(* Logix 5000 project; controller AOI_Working vendor 1 type 14 code 166 rev 35.11; software revision 35.04 *)

TASK MainTask (continuous, watchdog 500 ms) : MainProgram
TASK Normal_500ms (periodic, rate 500 ms, priority 10, watchdog 500 ms) : Main

MODULES
   Local : vendor 1 type 14 code 166 (ICP 0, rev 35.11)
END_MODULES

ADD_ON_INSTRUCTION AnalogInput   (* revision 1.1, vendor NixSoftware *)
// Simple scaling routine for analog inputs.
// Converts between raw units to EU
VAR_INPUT
   Inp_PVRaw : REAL; {required}   // Raw Input from I/O Point
   Cfg_InpRawMax : REAL := 100.0; {visible}   // Raw Value - Maximum Reading (Used for Scaling)
   Cfg_InpRawMin : REAL; {visible}   // Raw Value - Minimum Reading (Used for Scaling)
   Cfg_PVEUMax : REAL := 100.0; {visible}   // PV Maximum Value (In Engineering Units)
   Cfg_PVEUMin : REAL; {visible}   // PV Minimum Value (In Engineering Units)
END_VAR
VAR_OUTPUT
   Val_PV : REAL; {visible}   // Scaled PV (EU)
END_VAR
VAR_INPUT
   Sts_RangeError : BOOL;   // 1 = Range Invalid, Check Max/Mins
   Sts_CfgError : BOOL;   // 1 = Check Range, Protects against dividing by 0
END_VAR
VAR
   HMI_IOAssignment : STRING; {access None}
   HMI_Description : STRING; {access None}
   HMI_DisplayTag : STRING; {access None}
   _EUSpan : REAL; {access None}
   _RawSpan : REAL; {access None}
END_VAR

ROUTINE Logic   (* structured text *)
// Simple scaling routine for analog inputs.
// Converts between raw units to EU
   (* ============================================================
      Analog Input Scaling - Engineering Units Conversion
      Project  : Inavant Custom AOI Library
      AOI Name : AnalogInput
      ============================================================ *)
   
   (* --- Parameters / Tags (map to AOI InOut or UDT members) ---
      Inp_PVRaw       : REAL  - Raw analog input value (e.g. 0.0–32767.0 or 4.0–20.0 mA)
      Cfg_InpRawMin   : REAL  - Raw value corresponding to engineering minimum (e.g. 0.0 or 4.0)
      Cfg_InpRawMax   : REAL  - Raw value corresponding to engineering maximum (e.g. 32767.0 or 20.0)
      Cfg_EUMin       : REAL  - Engineering unit minimum (e.g. 0.0 PSI)
      Cfg_EUMax       : REAL  - Engineering unit maximum (e.g. 100.0 PSI)
      Val_PV         : REAL   - Scaled output in engineering units
      Sts_RangeErr    : BOOL  - Fault bit: TRUE if raw input is out of configured range
      Sts_DivZeroFlt  : BOOL  - Fault bit: TRUE if raw span is zero (invalid config)
   *)
   (* --- Clear faults from previous scan --- *)
   Sts_CfgError 		:= 0;
   Sts_RangeError   	:= 0;
   
   (* --- Guard: detect zero-span configuration --- *)
   _RawSpan := Cfg_InpRawMax - Cfg_InpRawMin;
   
   IF _RawSpan = 0.0 THEN
       (* Invalid config — cannot divide by zero; hold last good output *)
       Sts_CfgError := 1;
   
   ELSE
       (* --- Range check (informational, does NOT clamp output) --- *)
       IF (Inp_PVRaw < Cfg_InpRawMin) OR (Inp_PVRaw > Cfg_InpRawMax) THEN
           Sts_RangeError := 1;
       END_IF;
       (* --- Scaling equation --- *)
       Val_PV  := (Inp_PVRaw - Cfg_InpRawMin) * ((Cfg_PVEUMax - Cfg_PVEUMin) / (Cfg_InpRawMax - Cfg_InpRawMin)) + Cfg_PVEUMin;
   END_IF;
END_ROUTINE
END_ADD_ON_INSTRUCTION

ADD_ON_INSTRUCTION Inv_AI   (* revision 1.1, vendor NixSoftware *)
// Used for scaling a raw analog value to engineering units, includes alarm statuses and debounces.
VAR_INPUT
   Inp_PV : REAL; {visible}
   Inp_IOStatus : BOOL := 1; {visible}   // 1 = I/O Status is Good 0 = Alarm, generates Sts_Fail
   Inp_LoLoGate : BOOL := 1; {visible}   // 1 = Low-Low Sts Enabled
   Inp_LoGate : BOOL := 1; {visible}   // 1 = Low Sts Enabled
   Inp_HiGate : BOOL := 1; {visible}   // 1 = High Sts Enabled
   Inp_HiHiGate : BOOL := 1; {visible}   // 1 = High-High Sts Enabled
   Inp_FailGate : BOOL := 1; {visible}   // 1 = Fail Sts Enabled
   Cfg_InpRawMin : REAL; {visible}
   Cfg_InpRawMax : REAL := 100.0; {visible}
   Cfg_PVEUMin : REAL; {visible}
   Cfg_PVEUMax : REAL := 100.0; {visible}
   Cfg_HiHiLim : REAL := 1.5e+20;
   Cfg_HiHiDB : REAL := 1.0;
   Cfg_HiLim : REAL := 1.5e+20;
   Cfg_HiDB : REAL := 1.0;
   Cfg_LoLim : REAL := -1.5e+20;
   Cfg_LoDB : REAL := 1.0;
   Cfg_LoLoLim : REAL := -1.5e+20;
   Cfg_LoLoDB : REAL := 1.0;
   Cfg_FailHiLim : REAL := 104.0;   // PV (EU) High Fail Limit
   Cfg_FailLoLim : REAL := -3.0;   // PV (EU) Low Fail Limit
   Cfg_FailDB : REAL := 0.5;   // Failed PV DB
   Cfg_HiHiDlyOn : ALIAS FOR HiHi_Debounce.Cfg_DebounceON; {access None}
   Cfg_HiHiDlyOff : ALIAS FOR HiHi_Debounce.Cfg_DebounceOFF; {access None}
   Cfg_HiDlyOn : ALIAS FOR Hi_Debounce.Cfg_DebounceON; {access None}
   Cfg_HiDlyOff : ALIAS FOR Hi_Debounce.Cfg_DebounceOFF; {access None}
   Cfg_LoDlyOn : ALIAS FOR Lo_Debounce.Cfg_DebounceON; {access None}
   Cfg_LoDlyOff : ALIAS FOR Lo_Debounce.Cfg_DebounceOFF; {access None}
   Cfg_LoLoDlyOn : ALIAS FOR LoLo_Debounce.Cfg_DebounceON; {access None}
   Cfg_LoLoDlyOff : ALIAS FOR LoLo_Debounce.Cfg_DebounceOFF; {access None}
   Cfg_FailDlyOn : ALIAS FOR Fail_Debounce.Cfg_DebounceON; {access None}
   Cfg_FailDlyOff : ALIAS FOR Fail_Debounce.Cfg_DebounceOFF; {access None}
   Cfg_PVDecPlcs : INT := 2;
   Cfg_FiltTC : REAL;
END_VAR
VAR_OUTPUT
   Val : REAL; {access Read Only, visible}   // PV (EU)
   Sts_HiHi : BOOL; {visible}   // 1 = High-High Alarm Active
   Sts_Hi : BOOL; {visible}   // 1 = High Alarm Active
   Sts_Lo : BOOL; {visible}   // 1 = Low Alarm Active
   Sts_LoLo : BOOL; {visible}   // 1 = Low-Low Alarm Active
   Sts_Err : BOOL; {access Read Only, visible}   // 1 = Error in Configuration
   Sts_Fail : BOOL; {access Read Only, visible}   // 1 = Failed PV (Out of Range)
   Sts_FaultPresent : BOOL; {access Read Only}
   Val_Fault : DINT; {access Read Only}   // 0 = None 1 = Low Alm 2 = Hi Alm 3 = LoLo Alm 4 = HiHi Alm 32 = Failed PV 34 = Config. Error
   Val_PVEUMax : REAL; {access None, visible}
   Val_PVEUMin : REAL; {access None, visible}
END_VAR
VAR
   HMI_EU : STRING; {access None}
   HMI_Description : STRING; {access None}
   HMI_DisplayTag : STRING; {access None}
   HMI_Rack : STRING := 'RXXX'; {access None}
   HMI_Slot : STRING := 'SXX'; {access None}
   HMI_Channel : STRING := 'Ch.XX'; {access None}
   Wrk_InpDINT : DINT; {access None}
   Wrk_InpInfNaN : BOOL; {access None}
   Wrk_CalcedPV : REAL; {access None}   // Scaled Value - Pre Filtering
   Wrk_ScanT : TIMER := (PRE := 2147483647); {access None}
   HiHi_Debounce : Inv_Debounce; {access None}   // HiHi Alarm Debounce
   Wrk_HiHi : BOOL; {access None}   // Internal flag: High-High Status
   Hi_Debounce : Inv_Debounce; {access None}   // High Alarm Debounce
   Wrk_Hi : BOOL; {access None}   // Internal flag: High Status
   Wrk_Lo : BOOL; {access None}   // Internal flag: Lo Status
   Lo_Debounce : Inv_Debounce; {access None}   // Low Alarm Debounce
   Wrk_LoLo : BOOL; {access None}   // Internal Flag: Low-Low Status
   LoLo_Debounce : Inv_Debounce; {access None}   // Low-Low Alarm Debounce
   Wrk_Fault : DINT; {access None}   // Internal Fault Monitoring Tag
   Wrk_Fail : BOOL; {access None}   // Internal Flag: Fail Status
   Fail_Debounce : Inv_Debounce; {access None}   // Fail Alarm Debounce
   Wrk_Alpha : REAL;
   Wrk_FiltPV : REAL;
   Wrk_ScanTime : REAL;
   Wrk_UnfiltPV : REAL;
   Err_Raw : BOOL; {access Read Only}
   Err_EU : BOOL; {access Read Only}
   TempIOLocation : STRING; {access None}
END_VAR

ROUTINE Logic   (* ladder *)
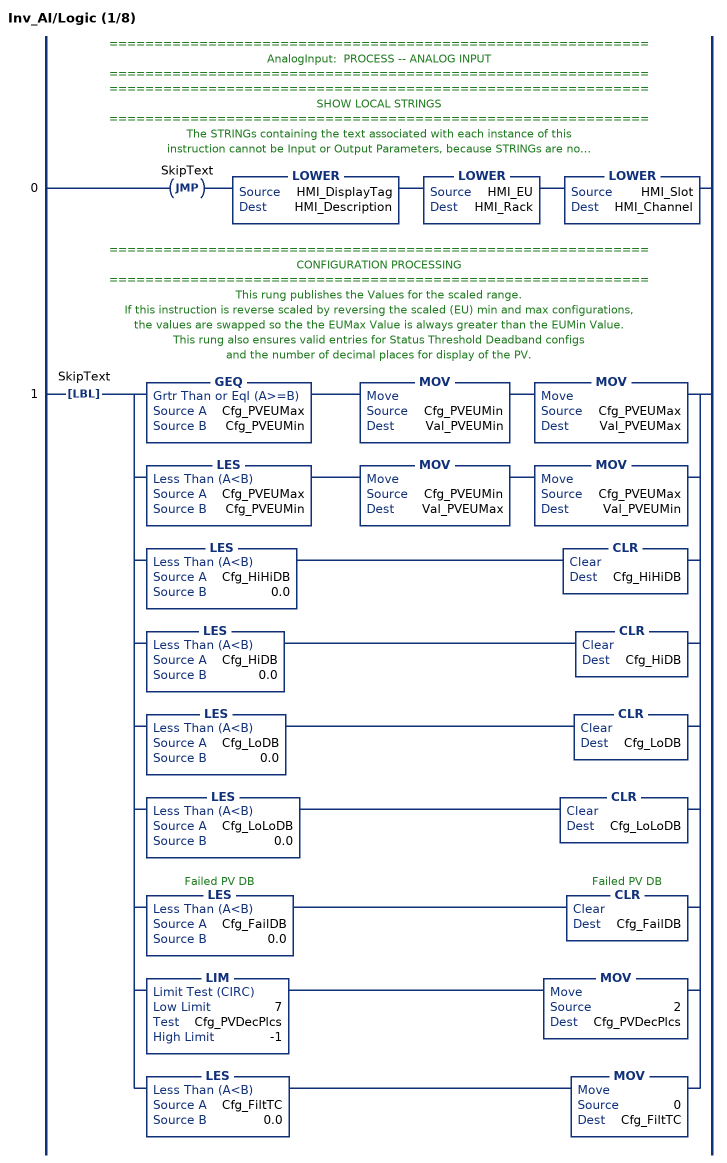
   // ============================================================
   // AnalogInput:  PROCESS -- ANALOG INPUT
   // ============================================================
   // ============================================================
   // SHOW LOCAL STRINGS
   // ============================================================
   // The STRINGs containing the text associated with each instance of this
   // instruction cannot be Input or Output Parameters, because STRINGs are not
   //  'atomic' types. (Inputs and Outputs must be SINT, INT, DINT, REAL, or BOOL.)
   // In order to make it easier to find and configure these STRINGs, this rung
   // was added.
   // Example as follows:
   // HMI_DisplayTag: FT-1234
   // HMI_Description: T-3 HCL Outfeed
   // HMI_EU: GPM
   // HMI_RACK: R150
   // HMI_Slot: S01
   // HMI_Channel: CH01
   0: JMP(SkipText)LOWER(HMI_DisplayTag,HMI_Description)LOWER(HMI_EU,HMI_Rack)LOWER(HMI_Slot,HMI_Channel);
   // ============================================================
   // CONFIGURATION PROCESSING
   // ============================================================
   // This rung publishes the Values for the scaled range.
   // If this instruction is reverse scaled by reversing the scaled (EU) min and max configurations,
   // the values are swapped so the the EUMax Value is always greater than the EUMin Value.
   // This rung also ensures valid entries for Status Threshold Deadband configs
   // and the number of decimal places for display of the PV.
   1: LBL(SkipText)[GEQ(Cfg_PVEUMax,Cfg_PVEUMin) MOV(Cfg_PVEUMin,Val_PVEUMin) MOV(Cfg_PVEUMax,Val_PVEUMax) ,LES(Cfg_PVEUMax,Cfg_PVEUMin) MOV(Cfg_PVEUMin,Val_PVEUMax) MOV(Cfg_PVEUMax,Val_PVEUMin) ,LES(Cfg_HiHiDB,0.0) CLR(Cfg_HiHiDB) ,LES(Cfg_HiDB,0.0) CLR(Cfg_HiDB) ,LES(Cfg_LoDB,0.0) CLR(Cfg_LoDB) ,LES(Cfg_LoLoDB,0.0) CLR(Cfg_LoLoDB) ,LES(Cfg_FailDB,0.0) CLR(Cfg_FailDB) ,LIM(7,Cfg_PVDecPlcs,-1) MOV(2,Cfg_PVDecPlcs) ,LES(Cfg_FiltTC,0.0) MOV(0,Cfg_FiltTC) ];
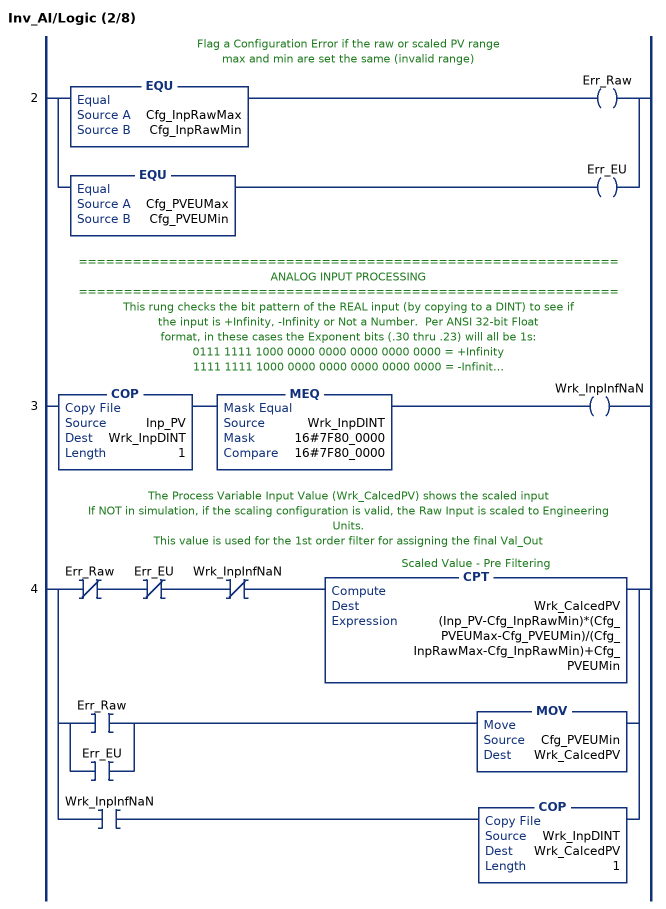
   // Flag a Configuration Error if the raw or scaled PV range
   // max and min are set the same (invalid range)
   2: [EQU(Cfg_InpRawMax,Cfg_InpRawMin) OTE(Err_Raw) ,EQU(Cfg_PVEUMax,Cfg_PVEUMin) OTE(Err_EU) ];
   // ============================================================
   // ANALOG INPUT PROCESSING
   // ============================================================
   // This rung checks the bit pattern of the REAL input (by copying to a DINT) to see if
   // the input is +Infinity, -Infinity or Not a Number.  Per ANSI 32-bit Float
   // format, in these cases the Exponent bits (.30 thru .23) will all be 1s:
   // 0111 1111 1000 0000 0000 0000 0000 0000 = +Infinity
   // 1111 1111 1000 0000 0000 0000 0000 0000 = -Infinity
   // x111 1111 1xxx xxxx xxxx xxxx xxxx xxxx = Not a Number
   3: COP(Inp_PV,Wrk_InpDINT,1)MEQ(Wrk_InpDINT,16#7F80_0000,16#7F80_0000)OTE(Wrk_InpInfNaN);
   // The Process Variable Input Value (Wrk_CalcedPV) shows the scaled input
   // If NOT in simulation, if the scaling configuration is valid, the Raw Input is scaled to Engineering Units.
   // This value is used for the 1st order filter for assigning the final Val_Out
   4: [XIO(Err_Raw) XIO(Err_EU) XIO(Wrk_InpInfNaN) CPT(Wrk_CalcedPV,(Inp_PV-Cfg_InpRawMin)*(Cfg_PVEUMax-Cfg_PVEUMin)/(Cfg_InpRawMax-Cfg_InpRawMin)+Cfg_PVEUMin) ,[XIC(Err_Raw) ,XIC(Err_EU) ] MOV(Cfg_PVEUMin,Wrk_CalcedPV) ,XIC(Wrk_InpInfNaN) COP(Wrk_InpDINT,Wrk_CalcedPV,1) ];
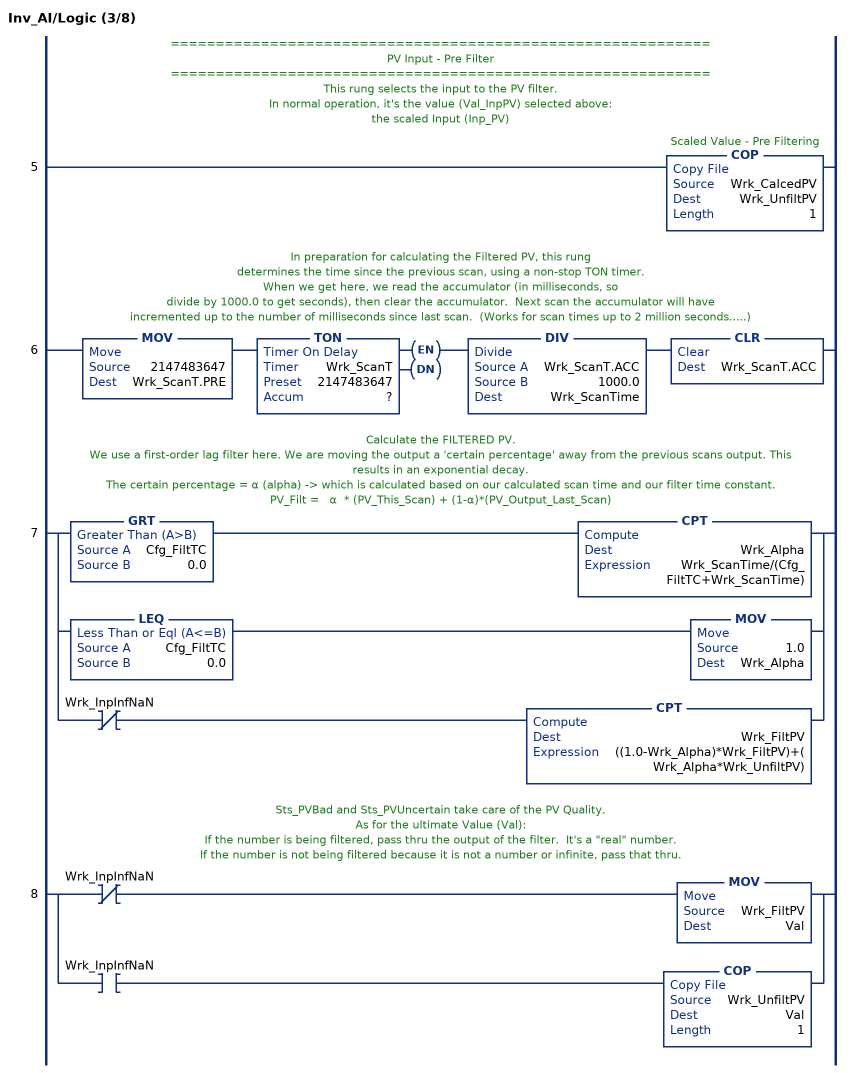
   // ============================================================
   // PV Input - Pre Filter
   // ============================================================
   // This rung selects the input to the PV filter.
   // In normal operation, it's the value (Val_InpPV) selected above:
   // the scaled Input (Inp_PV)
   5: COP(Wrk_CalcedPV,Wrk_UnfiltPV,1);
   // In preparation for calculating the Filtered PV, this rung
   // determines the time since the previous scan, using a non-stop TON timer.
   // When we get here, we read the accumulator (in milliseconds, so
   // divide by 1000.0 to get seconds), then clear the accumulator.  Next scan the accumulator will have
   // incremented up to the number of milliseconds since last scan.  (Works for scan times up to 2 million seconds.....)
   6: MOV(2147483647,Wrk_ScanT.PRE)TON(Wrk_ScanT,?,?)DIV(Wrk_ScanT.ACC,1000.0,Wrk_ScanTime)CLR(Wrk_ScanT.ACC);
   // Calculate the FILTERED PV.
   // We use a first-order lag filter here. We are moving the output a 'certain percentage' away from the previous scans output. This results in an exponential decay.
   // The certain percentage = α (alpha) -> which is calculated based on our calculated scan time and our filter time constant.
   // PV_Filt = 	α  * (PV_This_Scan) + (1-α)*(PV_Output_Last_Scan)
   7: [GRT(Cfg_FiltTC,0.0) CPT(Wrk_Alpha,Wrk_ScanTime/(Cfg_FiltTC+Wrk_ScanTime)) ,LEQ(Cfg_FiltTC,0.0) MOV(1.0,Wrk_Alpha) ,XIO(Wrk_InpInfNaN) CPT(Wrk_FiltPV,((1.0-Wrk_Alpha)*Wrk_FiltPV)+(Wrk_Alpha*Wrk_UnfiltPV)) ];
   // Sts_PVBad and Sts_PVUncertain take care of the PV Quality.
   // As for the ultimate Value (Val):
   // If the number is being filtered, pass thru the output of the filter.  It's a "real" number.
   // If the number is not being filtered because it is not a number or infinite, pass that thru.
   8: [XIO(Wrk_InpInfNaN) MOV(Wrk_FiltPV,Val) ,XIC(Wrk_InpInfNaN) COP(Wrk_UnfiltPV,Val,1) ];
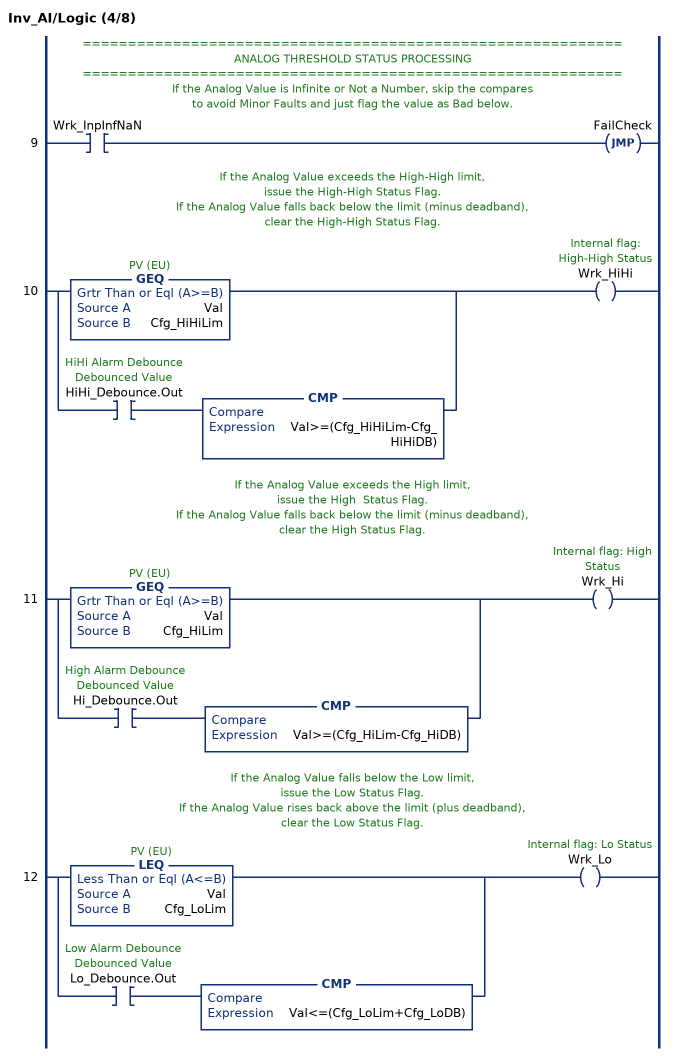
   // ============================================================
   // ANALOG THRESHOLD STATUS PROCESSING
   // ============================================================
   // If the Analog Value is Infinite or Not a Number, skip the compares
   // to avoid Minor Faults and just flag the value as Bad below.
   9: XIC(Wrk_InpInfNaN)JMP(FailCheck);
   // If the Analog Value exceeds the High-High limit,
   // issue the High-High Status Flag.
   // If the Analog Value falls back below the limit (minus deadband),
   // clear the High-High Status Flag.
   10: [GEQ(Val,Cfg_HiHiLim) ,XIC(HiHi_Debounce.Out) CMP(Val>=(Cfg_HiHiLim-Cfg_HiHiDB)) ]OTE(Wrk_HiHi);
   // If the Analog Value exceeds the High limit,
   // issue the High  Status Flag.
   // If the Analog Value falls back below the limit (minus deadband),
   // clear the High Status Flag.
   11: [GEQ(Val,Cfg_HiLim) ,XIC(Hi_Debounce.Out) CMP(Val>=(Cfg_HiLim-Cfg_HiDB)) ]OTE(Wrk_Hi);
   // If the Analog Value falls below the Low limit,
   // issue the Low Status Flag.
   // If the Analog Value rises back above the limit (plus deadband),
   // clear the Low Status Flag.
   12: [LEQ(Val,Cfg_LoLim) ,XIC(Lo_Debounce.Out) CMP(Val<=(Cfg_LoLim+Cfg_LoDB)) ]OTE(Wrk_Lo);
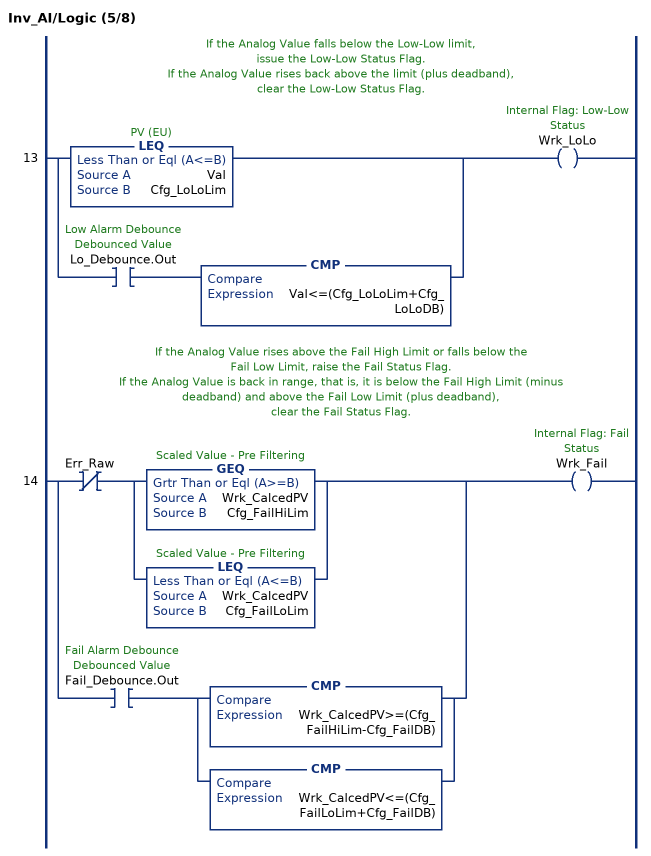
   // If the Analog Value falls below the Low-Low limit,
   // issue the Low-Low Status Flag.
   // If the Analog Value rises back above the limit (plus deadband),
   // clear the Low-Low Status Flag.
   13: [LEQ(Val,Cfg_LoLoLim) ,XIC(Lo_Debounce.Out) CMP(Val<=(Cfg_LoLoLim+Cfg_LoLoDB)) ]OTE(Wrk_LoLo);
   // If the Analog Value rises above the Fail High Limit or falls below the
   // Fail Low Limit, raise the Fail Status Flag.
   // If the Analog Value is back in range, that is, it is below the Fail High Limit (minus
   // deadband) and above the Fail Low Limit (plus deadband),
   // clear the Fail Status Flag.
   14: [XIO(Err_Raw) [GEQ(Wrk_CalcedPV,Cfg_FailHiLim) ,LEQ(Wrk_CalcedPV,Cfg_FailLoLim) ] ,XIC(Fail_Debounce.Out) [CMP(Wrk_CalcedPV>=(Cfg_FailHiLim-Cfg_FailDB)) ,CMP(Wrk_CalcedPV<=(Cfg_FailLoLim+Cfg_FailDB)) ] ]OTE(Wrk_Fail);
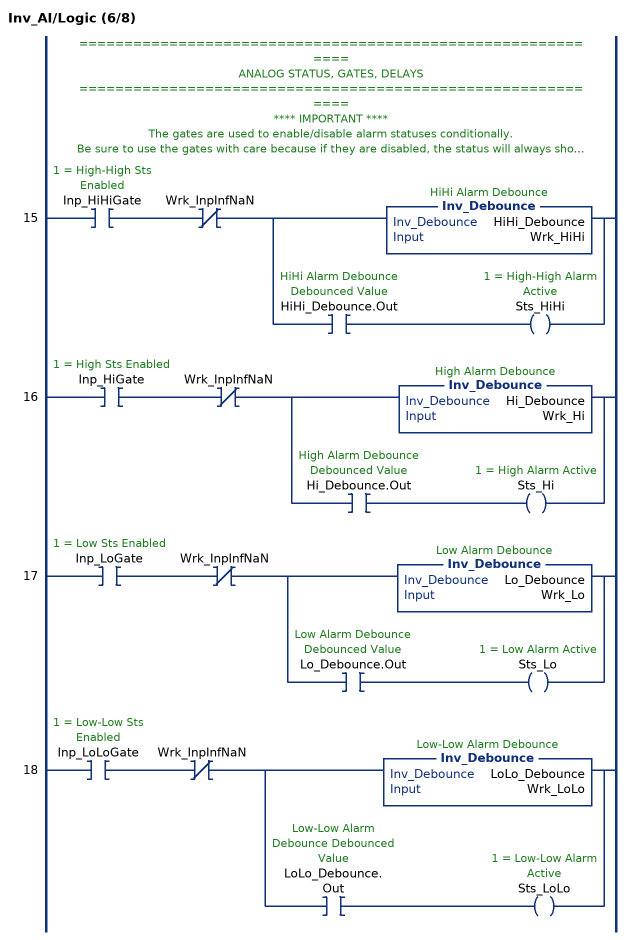
   // ============================================================
   // ANALOG STATUS, GATES, DELAYS
   // ============================================================
   // **** IMPORTANT ****
   // The gates are used to enable/disable alarm statuses conditionally.
   // Be sure to use the gates with care because if they are disabled, the status will always show off.
   15: XIC(Inp_HiHiGate)XIO(Wrk_InpInfNaN)[Inv_Debounce(HiHi_Debounce,Wrk_HiHi) ,XIC(HiHi_Debounce.Out) OTE(Sts_HiHi) ];
   16: XIC(Inp_HiGate)XIO(Wrk_InpInfNaN)[Inv_Debounce(Hi_Debounce,Wrk_Hi) ,XIC(Hi_Debounce.Out) OTE(Sts_Hi) ];
   17: XIC(Inp_LoGate)XIO(Wrk_InpInfNaN)[Inv_Debounce(Lo_Debounce,Wrk_Lo) ,XIC(Lo_Debounce.Out) OTE(Sts_Lo) ];
   18: XIC(Inp_LoLoGate)XIO(Wrk_InpInfNaN)[Inv_Debounce(LoLo_Debounce,Wrk_LoLo) ,XIC(LoLo_Debounce.Out) OTE(Sts_LoLo) ];
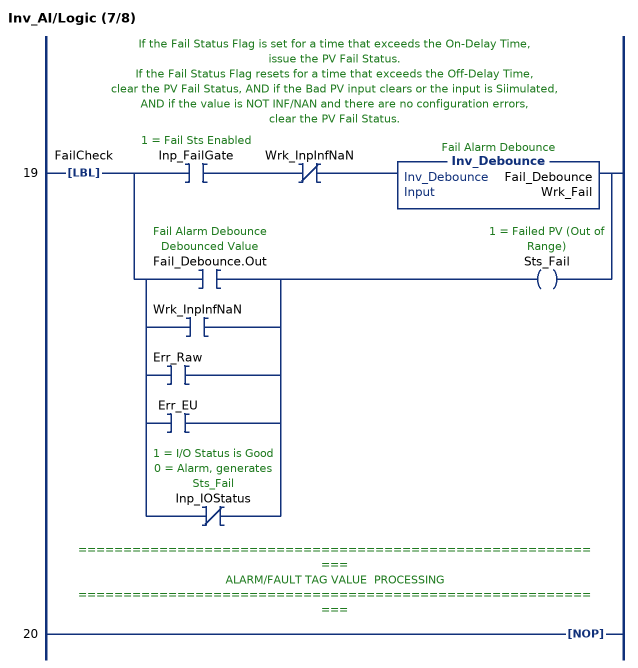
   // If the Fail Status Flag is set for a time that exceeds the On-Delay Time,
   // issue the PV Fail Status.
   // If the Fail Status Flag resets for a time that exceeds the Off-Delay Time,
   // clear the PV Fail Status, AND if the Bad PV input clears or the input is Siimulated,
   // AND if the value is NOT INF/NAN and there are no configuration errors,
   // clear the PV Fail Status.
   19: LBL(FailCheck)[XIC(Inp_FailGate) XIO(Wrk_InpInfNaN) Inv_Debounce(Fail_Debounce,Wrk_Fail) ,[XIC(Fail_Debounce.Out) ,XIC(Wrk_InpInfNaN) ,XIC(Err_Raw) ,XIC(Err_EU) ,XIO(Inp_IOStatus) ] OTE(Sts_Fail) ];
   // ============================================================
   // ALARM/FAULT TAG VALUE  PROCESSING
   // ============================================================
   20: NOP();
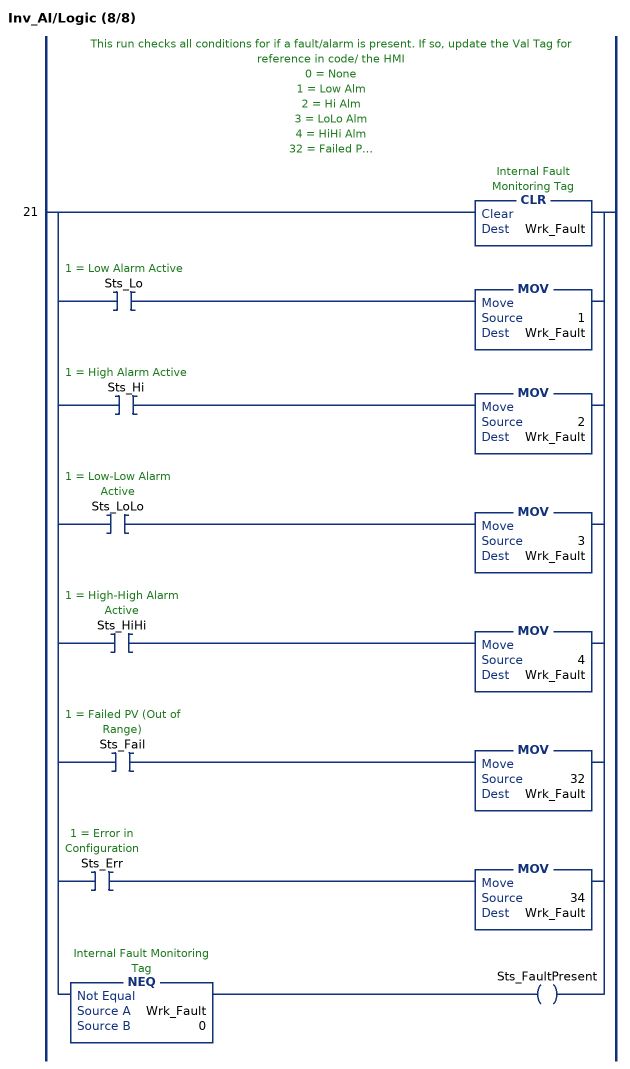
   // This run checks all conditions for if a fault/alarm is present. If so, update the Val Tag for reference in code/ the HMI
   // 0 = None
   // 1 = Low Alm
   // 2 = Hi Alm
   // 3 = LoLo Alm
   // 4 = HiHi Alm
   // 32 = Failed PV
   // 34 = Config. Error
   21: [CLR(Wrk_Fault) ,XIC(Sts_Lo) MOV(1,Wrk_Fault) ,XIC(Sts_Hi) MOV(2,Wrk_Fault) ,XIC(Sts_LoLo) MOV(3,Wrk_Fault) ,XIC(Sts_HiHi) MOV(4,Wrk_Fault) ,XIC(Sts_Fail) MOV(32,Wrk_Fault) ,XIC(Sts_Err) MOV(34,Wrk_Fault) ,NEQ(Wrk_Fault,0) OTE(Sts_FaultPresent) ];
END_ROUTINE
END_ADD_ON_INSTRUCTION

ADD_ON_INSTRUCTION Inv_Debounce   (* revision 1.1, vendor NixSoftware *)
// Can be dropped into any ladder routine on its own and used to debounce a discrete input.
// Assign the input channel or alias to 'Input' and use the .Out value anywhere the DI would be used instead.
VAR_INPUT
   Input : BOOL; {required}   // Raw Input to be debounced
   Cfg_DebounceON : REAL; {visible}   // Time (s) to debounce input before turning Out status ON Range (0-30s)
   Cfg_DebounceOFF : REAL; {visible}   // Time (s) to debounce input before turning Out status OFF Range (0-30s)
END_VAR
VAR_OUTPUT
   Out : BOOL; {access Read Only, visible}   // Debounced Value
END_VAR
VAR
   DebounceMaxTime : REAL := 30.0; {access None}
   Work_RiseT : TIMER; {access None}
   Work_FallT : TIMER; {access None}
END_VAR

ROUTINE Logic   (* ladder *)
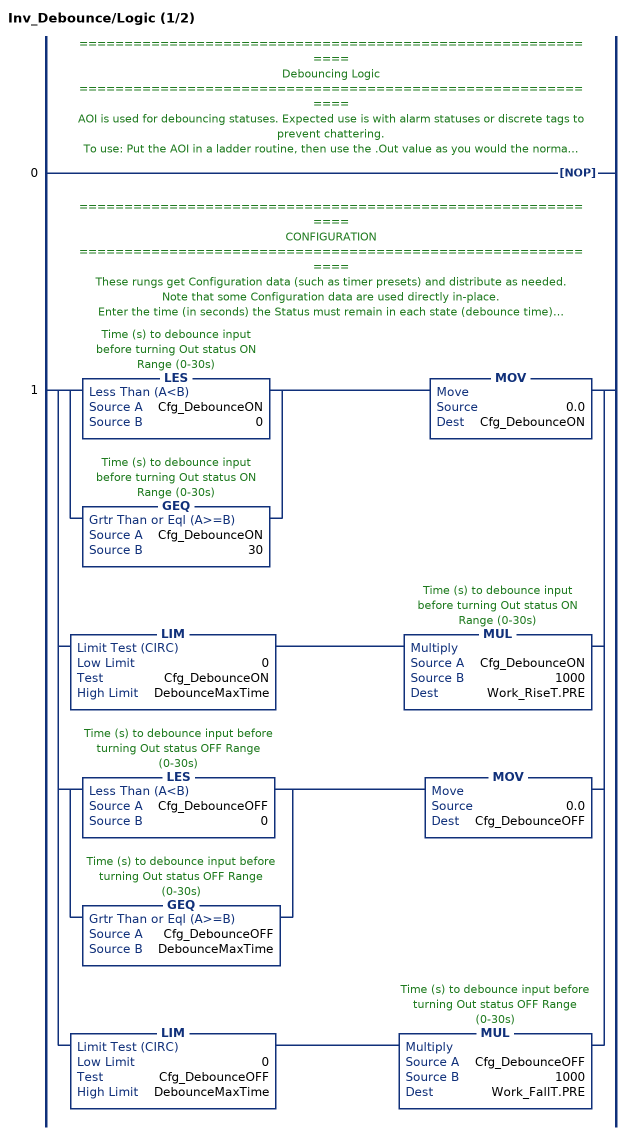
   // ============================================================
   // Debouncing Logic
   // ============================================================
   // AOI is used for debouncing statuses. Expected use is with alarm statuses or discrete tags to prevent chattering.
   // To use: Put the AOI in a ladder routine, then use the .Out value as you would the normal input to use the debounced value.
   0: NOP();
   // ============================================================
   // CONFIGURATION
   // ============================================================
   // These rungs get Configuration data (such as timer presets) and distribute as needed.
   // Note that some Configuration data are used directly in-place.
   // Enter the time (in seconds) the Status must remain in each state (debounce time).
   // There is a time used for the rising-edge and falling-edge debounce
   // If our Debounce time preset is out of range (Negative or greater than MaxDebounce) -> Move a 0 to the value to prevent a major controller fault on a negative timer preset
   1: [[LES(Cfg_DebounceON,0) ,GEQ(Cfg_DebounceON,30) ] MOV(0.0,Cfg_DebounceON) ,LIM(0,Cfg_DebounceON,DebounceMaxTime) MUL(Cfg_DebounceON,1000,Work_RiseT.PRE) ,[LES(Cfg_DebounceOFF,0) ,GEQ(Cfg_DebounceOFF,DebounceMaxTime) ] MOV(0.0,Cfg_DebounceOFF) ,LIM(0,Cfg_DebounceOFF,DebounceMaxTime) MUL(Cfg_DebounceOFF,1000,Work_FallT.PRE) ];
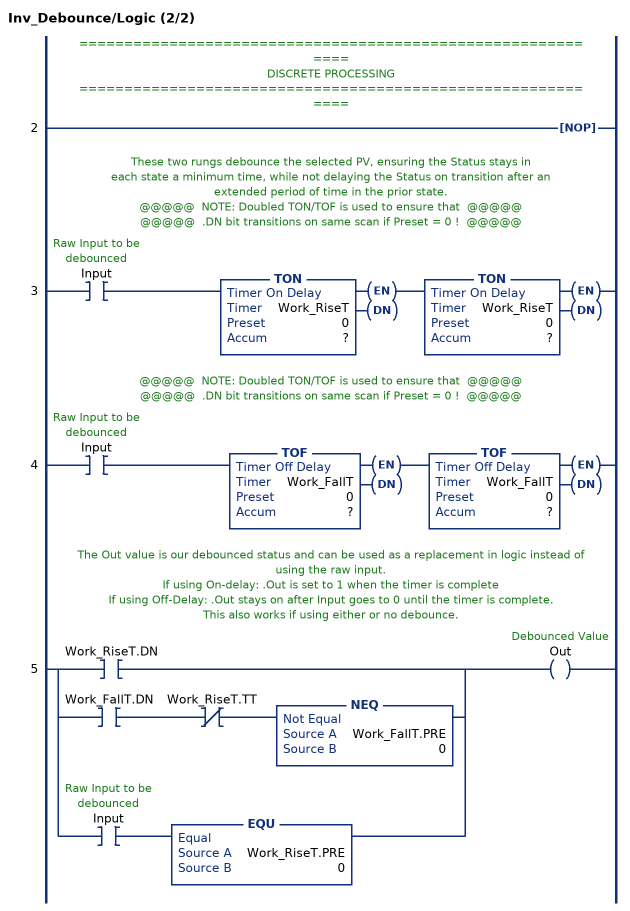
   // ============================================================
   // DISCRETE PROCESSING
   // ============================================================
   2: NOP();
   // These two rungs debounce the selected PV, ensuring the Status stays in
   // each state a minimum time, while not delaying the Status on transition after an
   // extended period of time in the prior state.
   // @@@@@  NOTE: Doubled TON/TOF is used to ensure that  @@@@@
   // @@@@@  .DN bit transitions on same scan if Preset = 0 !  @@@@@
   3: XIC(Input)TON(Work_RiseT,?,?)TON(Work_RiseT,?,?);
   // @@@@@  NOTE: Doubled TON/TOF is used to ensure that  @@@@@
   // @@@@@  .DN bit transitions on same scan if Preset = 0 !  @@@@@
   4: XIC(Input)TOF(Work_FallT,?,?)TOF(Work_FallT,?,?);
   // The Out value is our debounced status and can be used as a replacement in logic instead of
   // using the raw input.
   // If using On-delay: .Out is set to 1 when the timer is complete
   // If using Off-Delay: .Out stays on after Input goes to 0 until the timer is complete.
   // This also works if using either or no debounce.
   5: [XIC(Work_RiseT.DN) ,XIC(Work_FallT.DN) XIO(Work_RiseT.TT) NEQ(Work_FallT.PRE,0) ,XIC(Input) EQU(Work_RiseT.PRE,0) ]OTE(Out);
END_ROUTINE
END_ADD_ON_INSTRUCTION

ADD_ON_INSTRUCTION Inv_FVNR   (* revision 1.0, vendor Inavant *)
// AOI for Non-Reversing Motor Starter
VAR_INPUT
   Cmd_Auto : BOOL;   // 1 = Auto 0 = Manual
END_VAR
VAR_OUTPUT
   Out_Run : BOOL; {access Read Only, required}
END_VAR
VAR_INPUT
   Inp_RunFdbk : BOOL; {required}
   Inp_ReadyStatus : BOOL; {required}   // Motor Ready Status ( 1 = Good ) (0 = Not Ready)
   Inp_IO_Ok : BOOL := 1; {visible}   // 1 = Good Comms 0 = Fault
   Intlk_OK : BOOL := 1; {visible}
   AutoCmd_Start : BOOL; {visible}   // Automatic Start Command
   AutoCmd_Stop : BOOL; {visible}   // Automatic Stop Command
   PBCmd_Start : BOOL; {visible}   // 1 = Local Start PB Cmd
   PBCmd_Stop : BOOL; {visible}   // 1 = Local Stop PB Cmd
END_VAR
VAR_OUTPUT
   Flt_Comm : BOOL; {access Read Only, visible}   // 1 = Comm. Fault, Check Device
   Flt_FailToStart : BOOL; {access Read Only, visible}
   Flt_FailToStop : BOOL; {access Read Only, visible}
   Flt_DeviceNotRdy : BOOL; {visible}
   Flt_MotorNotReady : BOOL; {access Read Only, visible}   // 1 = Motor Not Ready to Run (Check Motor Bucket)
   Sts_Auto : BOOL := 1; {visible}
   Sts_Manual : BOOL;
END_VAR
VAR_INPUT
   AutoCmd_ResetFaults : BOOL; {visible}
   Cfg_EnFailToStartFlt : BOOL := 1;   // 1 = Enable Fail to Start Fault
   Cfg_EnFailToStopFlt : BOOL := 1;
   Cfg_EnCommsFlt : BOOL := 1;
   Cfg_EnDeviceNotRdyFlt : BOOL := 1;   // 1 = Enable Fail to Start Fault
   Cfg_UseRunFdbk : BOOL := 1;
   Cfg_FTStOrStpPRE : REAL := 10.0;   // Time (s) for the Fai to Start or Stop Timer (0-30s)
END_VAR
VAR_OUTPUT
   Val_Sts : DINT; {visible}   // 0 = STOPPED 1 = STARTING 2 = RUNNING 3 = STOPPING
END_VAR
VAR_INPUT
   Sts_Faulted : BOOL; {visible}
   Val_Fault : DINT;   // 0 = Good, No Faults 1 = Fail To Start 2 = Fail To Stop 5 = Comm/IO Fault
   Cmd_ResetFaults : BOOL;
   Cfg_EnMotorRdyFlt : BOOL := 1;
END_VAR
VAR_OUTPUT
   Sts_Running : BOOL; {access Read Only, visible}
   Sts_Ready2Run : BOOL; {access Read Only, visible}   // Motor has no faults and isn't interlocked - Ready to Run
END_VAR
VAR
   TMR_FlToStOrStp : TIMER := (PRE := 7000); {access None}
   TMR_MinHoldReset : TIMER := (PRE := 1000); {access None}   // Minimum Reset Pulse Time
   TMR_HoldReset : TIMER := (PRE := 1000); {access None}   // Timer that sets Maximum Reset Pulse Time based on how long Operator is pressing button
   HMI_Cmd_Reset : BOOL;
   HMI_Cmd_Stop : BOOL;
   HMI_Cmd_Start : BOOL;
   Wrk_RunDwn : BOOL; {access None}
   Wrk_RunUp : BOOL; {access None}
END_VAR

ROUTINE Logic   (* ladder *)
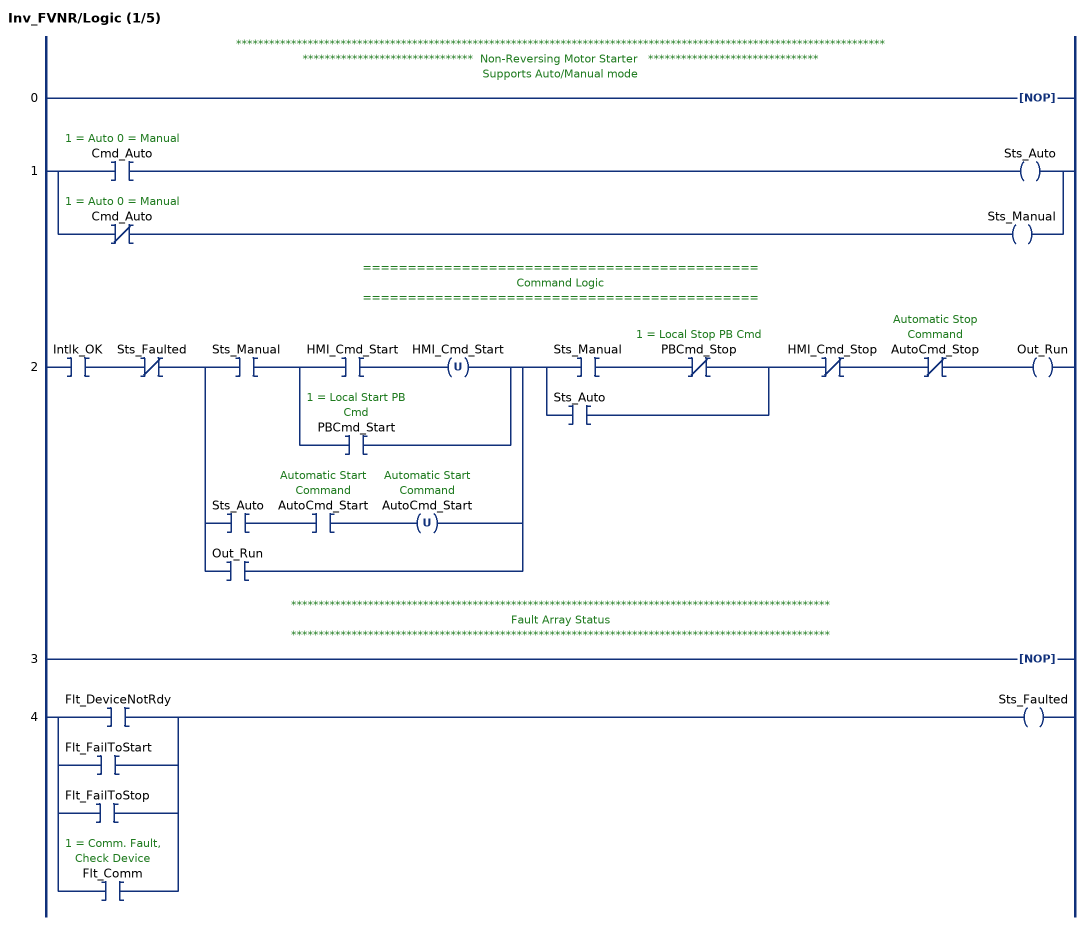
   // **********************************************************************************************************************
   // *******************************  Non-Reversing Motor Starter   *******************************
   // Supports Auto/Manual mode
   0: NOP();
   1: [XIC(Cmd_Auto) OTE(Sts_Auto) ,XIO(Cmd_Auto) OTE(Sts_Manual) ];
   // ============================================
   // Command Logic
   // ============================================
   2: XIC(Intlk_OK)XIO(Sts_Faulted)[XIC(Sts_Manual) [XIC(HMI_Cmd_Start) OTU(HMI_Cmd_Start) ,XIC(PBCmd_Start) ] ,XIC(Sts_Auto) XIC(AutoCmd_Start) OTU(AutoCmd_Start) ,XIC(Out_Run) ][XIC(Sts_Manual) XIO(PBCmd_Stop) ,XIC(Sts_Auto) ]XIO(HMI_Cmd_Stop)XIO(AutoCmd_Stop)OTE(Out_Run);
   // **************************************************************************************************
   // Fault Array Status
   // **************************************************************************************************
   3: NOP();
   4: [XIC(Flt_DeviceNotRdy) ,XIC(Flt_FailToStart) ,XIC(Flt_FailToStop) ,XIC(Flt_Comm) ]OTE(Sts_Faulted);
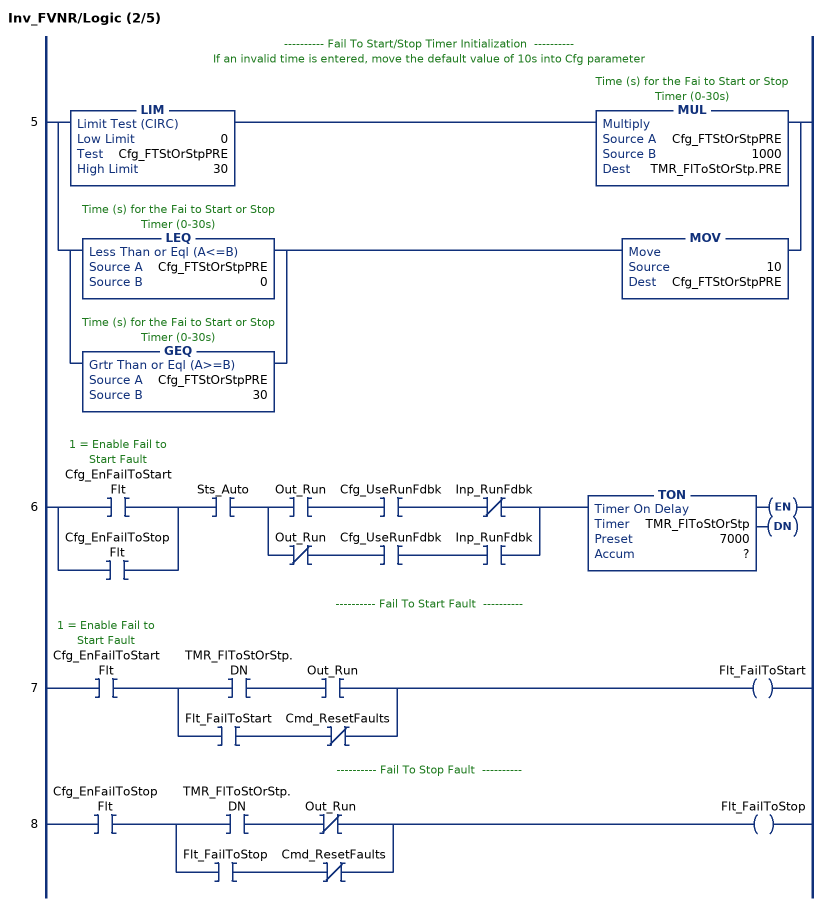
   // ---------- Fail To Start/Stop Timer Initialization  ----------
   // If an invalid time is entered, move the default value of 10s into Cfg parameter
   5: [LIM(0,Cfg_FTStOrStpPRE,30) MUL(Cfg_FTStOrStpPRE,1000,TMR_FlToStOrStp.PRE) ,[LEQ(Cfg_FTStOrStpPRE,0) ,GEQ(Cfg_FTStOrStpPRE,30) ] MOV(10,Cfg_FTStOrStpPRE) ];
   6: [XIC(Cfg_EnFailToStartFlt) ,XIC(Cfg_EnFailToStopFlt) ]XIC(Sts_Auto)[XIC(Out_Run) XIC(Cfg_UseRunFdbk) XIO(Inp_RunFdbk) ,XIO(Out_Run) XIC(Cfg_UseRunFdbk) XIC(Inp_RunFdbk) ]TON(TMR_FlToStOrStp,?,?);
   // ---------- Fail To Start Fault  ----------
   7: XIC(Cfg_EnFailToStartFlt)[XIC(TMR_FlToStOrStp.DN) XIC(Out_Run) ,XIC(Flt_FailToStart) XIO(Cmd_ResetFaults) ]OTE(Flt_FailToStart);
   // ---------- Fail To Stop Fault  ----------
   8: XIC(Cfg_EnFailToStopFlt)[XIC(TMR_FlToStOrStp.DN) XIO(Out_Run) ,XIC(Flt_FailToStop) XIO(Cmd_ResetFaults) ]OTE(Flt_FailToStop);
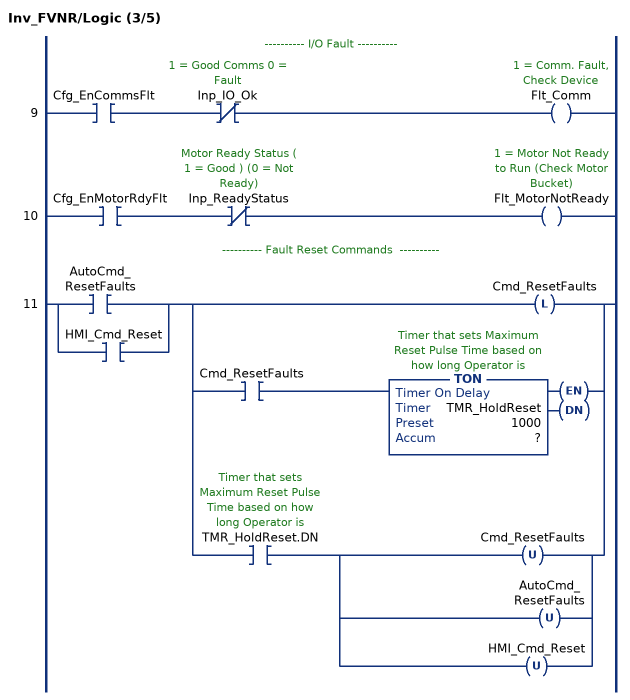
   // ---------- I/O Fault ----------
   9: XIC(Cfg_EnCommsFlt)XIO(Inp_IO_Ok)OTE(Flt_Comm);
   10: XIC(Cfg_EnMotorRdyFlt)XIO(Inp_ReadyStatus)OTE(Flt_MotorNotReady);
   // ---------- Fault Reset Commands  ----------
   11: [XIC(AutoCmd_ResetFaults) ,XIC(HMI_Cmd_Reset) ][OTL(Cmd_ResetFaults) ,XIC(Cmd_ResetFaults) TON(TMR_HoldReset,?,?) ,XIC(TMR_HoldReset.DN) [OTU(Cmd_ResetFaults) ,OTU(AutoCmd_ResetFaults) ,OTU(HMI_Cmd_Reset) ] ];
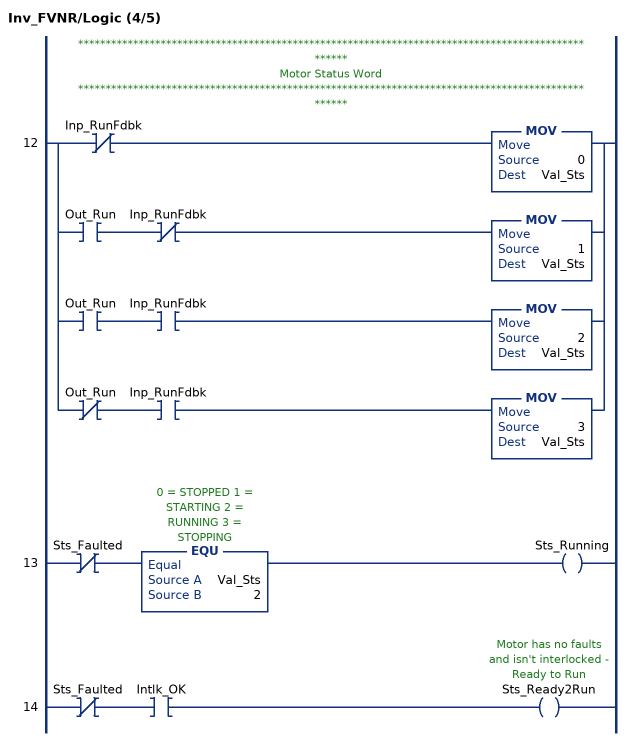
   // **************************************************************************************************
   // Motor Status Word
   // **************************************************************************************************
   12: [XIO(Inp_RunFdbk) MOV(0,Val_Sts) ,XIC(Out_Run) XIO(Inp_RunFdbk) MOV(1,Val_Sts) ,XIC(Out_Run) XIC(Inp_RunFdbk) MOV(2,Val_Sts) ,XIO(Out_Run) XIC(Inp_RunFdbk) MOV(3,Val_Sts) ];
   13: XIO(Sts_Faulted)EQU(Val_Sts,2)OTE(Sts_Running);
   14: XIO(Sts_Faulted)XIC(Intlk_OK)OTE(Sts_Ready2Run);
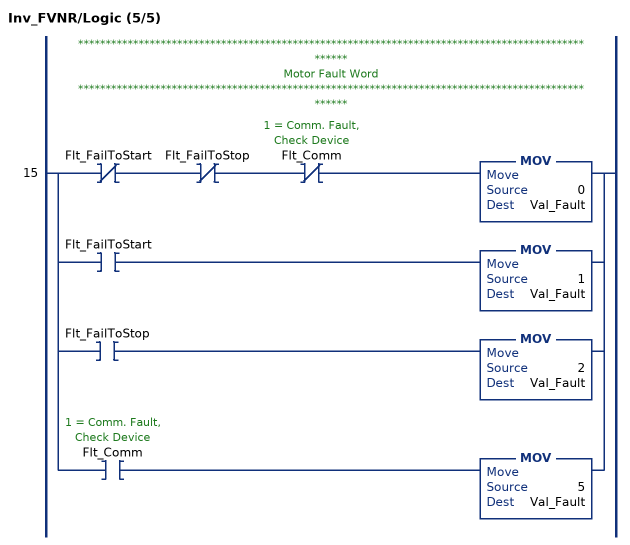
   // **************************************************************************************************
   // Motor Fault Word
   // **************************************************************************************************
   15: [XIO(Flt_FailToStart) XIO(Flt_FailToStop) XIO(Flt_Comm) MOV(0,Val_Fault) ,XIC(Flt_FailToStart) MOV(1,Val_Fault) ,XIC(Flt_FailToStop) MOV(2,Val_Fault) ,XIC(Flt_Comm) MOV(5,Val_Fault) ];
END_ROUTINE
END_ADD_ON_INSTRUCTION

ADD_ON_INSTRUCTION Inv_ModuleStatus   (* revision 1.1 *)
// I/O Status
VAR_IN_OUT
   ModuleName : MODULE; {required}
END_VAR
VAR_INPUT
   Inp_Sim : BOOL;
   Set_SimFault : BOOL;
END_VAR
VAR_OUTPUT
   Sts_IOFault : BOOL; {access Read Only, visible}
   Val_Fault : DINT; {access Read Only, visible}
END_VAR
VAR
   EntrySts : INT; {access None}
   ConnectionSts : DINT; {access None}
   FaultVal : DINT; {access None}
END_VAR

ROUTINE Logic   (* ladder *)
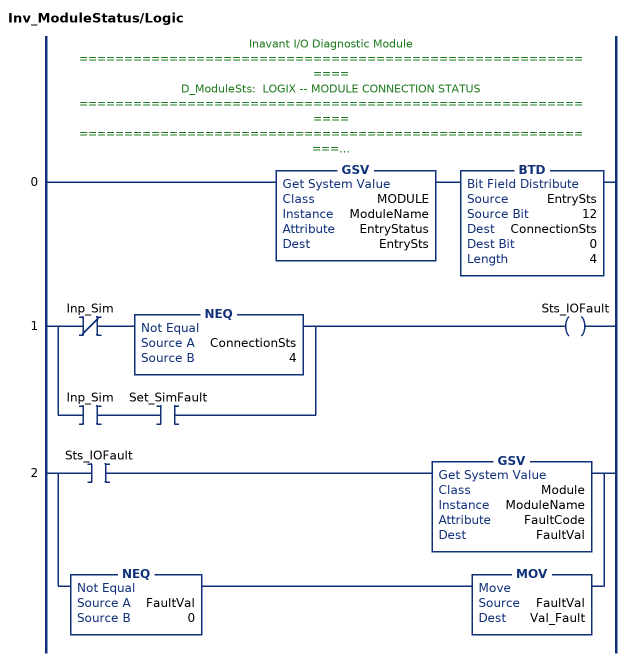
   // Inavant I/O Diagnostic Module
   // ============================================================
   // D_ModuleSts:  LOGIX -- MODULE CONNECTION STATUS
   // ============================================================
   // ============================================================
   // This Instruction monitors the connection status of one Module
   // in the Logix controller's I/O Configuration tree and provides
   // an I/O Fault status if the connection is NOT "Running".
   // ============================================================
   // Use a GSV to the MODULE object to get the "EntryStatus" attribute.
   0: GSV(MODULE,ModuleName,EntryStatus,EntrySts)BTD(EntrySts,12,ConnectionSts,0,4);
   1: [XIO(Inp_Sim) NEQ(ConnectionSts,4) ,XIC(Inp_Sim) XIC(Set_SimFault) ]OTE(Sts_IOFault);
   2: [XIC(Sts_IOFault) GSV(Module,ModuleName,FaultCode,FaultVal) ,NEQ(FaultVal,0) MOV(FaultVal,Val_Fault) ];
END_ROUTINE
END_ADD_ON_INSTRUCTION

VAR_GLOBAL   (* controller tags *)
   AI_Test : AnalogInput := (Cfg_InpRawMax := 100.0, Cfg_PVEUMax := 100.0);
   AI_Test2 : AnalogInput := (Cfg_InpRawMax := 100.0, Cfg_PVEUMax := 100.0);
   PT_1234 : REAL;
END_VAR

PROGRAM Main   (* main routine AnalogInputTest *)
VAR
   AI_Test1 : AnalogInput := (Cfg_InpRawMax := 100.0, Cfg_PVEUMax := 100.0);
   SCL_01 : SCALE;
END_VAR

ROUTINE AnalogInputFBD   (* function block diagram *)
   SHEET 1
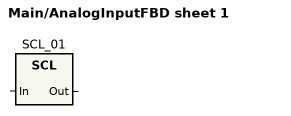
   SCL_01 : SCL();   // unwired pins: In Out
END_ROUTINE

ROUTINE AnalogInputTest   (* ladder *)
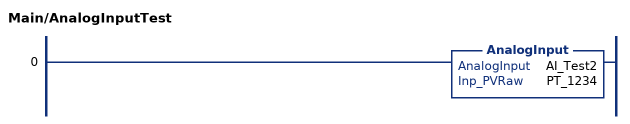
   0: AnalogInput(AI_Test2,PT_1234);
END_ROUTINE
END_PROGRAM

PROGRAM MainProgram   (* main routine MainRoutine *)

ROUTINE MainRoutine   (* ladder *)
END_ROUTINE
END_PROGRAM
